// TIA Portal V21 export
// export: Created 2026-11-11T00:48:23.7852385Z, ExportSetting WithDefaults, DisplayName Totally Integrated Automation Portal, DisplayVersion V21 Update 3, DisplayName STEP 7 Professional, DisplayVersion V21 Update 3, DisplayName STEP 7 Safety, DisplayVersion V21, DisplayName Tech WebApplication, DisplayVersion V21, DisplayName WinCC Basic/Comfort/Advanced, DisplayVersion V21 Update 3, DisplayName WinCC Unified, DisplayVersion V21 Update 3
FUNCTION_BLOCK "FB_Scl_sl114"   // FB198, SCL
{ S7_Optimized_Access := 'TRUE' }
VERSION : 0.1
// stored: AutoNumber true, IsIECCheckEnabled false, IsRetainMemResEnabled false, MemoryReserve 100, SetENOAutomatically false, UDAEnableTagReadback false
   VAR_INPUT
      v_o_cmd : Bool;
      v_c_cmd : Bool;
      v_s_cmd : Bool;
      v_o_fb : Bool;
      v_c_fb : Bool;
   END_VAR
   VAR_OUTPUT
      v_oo : Bool;
      v_co : Bool;
      v_oa : Bool;
      v_ca : Bool;
      v_q : Bool;
   END_VAR
   VAR
      inst { S7_SetPoint := 'True'} : MCAT;
   END_VAR
BEGIN
   #inst(O_CMD := #v_o_cmd, C_CMD := #v_c_cmd, S_CMD := #v_s_cmd, O_FB := #v_o_fb, C_FB := #v_c_fb, OO => #v_oo, CO => #v_co, OA => #v_oa, CA => #v_ca, Q => #v_q);
END_FUNCTION_BLOCK
